TYPE ST_WeldingStatus :
STRUCT
	lrStartWelding				:LREAL;
	lrEndWelding					:LREAL;
	lrDistanceWelding				:LREAL;
END_STRUCT
END_TYPE

(* stored: Version 1.1.0.1, ProductVersion 3.1.4024.15
   DUT ST_WeldingStatus: Id {ecd4be42-75d3-439f-ba6a-57d0692f3c97} *)
